(* CODESYS project Example8_PLC.project

Project tree, tasks and I/O mapping:
  Device : CODESYS Control Win V3, 3S - Smart Software Solutions GmbH, order no. 305021, version 3.5.7.0
    application Application
      libraries: Standard, * (System)
      task MainTask (cyclic, interval t#20ms, priority 1) calls PLC_PRG
      program PLC_PRG [ST]
      global variables GVL
      function block FB_G4LTL [ST]
    Ethernet : Ethernet, 3S - Smart Software Solutions GmbH, version 3.5.7.0
      Modbus_TCP_Master : Modbus TCP Master, 3S - Smart Software Solutions GmbH, version 3.5.6.0
          settings: AutoReconnect = TRUE
        Modbus_TCP_Slave : Modbus TCP Slave, 3S - Smart Software Solutions GmbH, version 3.5.7.0
            settings: Unit-ID = 1; IPAddress = [127, 0, 0, 1]; Channel 0.Function Code = 4; Channel 0.Read Offset = 16#0000; Channel 0.Read Length = 1; Channel 0.Write Offset = 0; Channel 0.Write Length = 0; Channel 0.Cycle Time = 100; Channel 1.Function Code = 4; Channel 1.Read Offset = 16#0001; Channel 1.Read Length = 1; Channel 1.Write Offset = 0; Channel 1.Write Length = 0; Channel 1.Cycle Time = 100; Channel 2.Function Code = 4; Channel 2.Read Offset = 16#0002; Channel 2.Read Length = 1; Channel 2.Write Offset = 0; Channel 2.Write Length = 0; Channel 2.Cycle Time = 100; Channel 3.Function Code = 4; Channel 3.Read Offset = 16#0003; Channel 3.Read Length = 1; Channel 3.Write Offset = 0; Channel 3.Write Length = 0; Channel 3.Cycle Time = 100; Channel 4.Function Code = 4; Channel 4.Read Offset = 16#0004; Channel 4.Read Length = 1; Channel 4.Write Offset = 0; Channel 4.Write Length = 0; Channel 4.Cycle Time = 100; Channel 5.Function Code = 6; Channel 5.Read Offset = 0; Channel 5.Read Length = 0; Channel 5.Write Offset = 16#0000; Channel 5.Write Length = 1; Channel 5.Cycle Time = 100; Channel 6.Function Code = 6; Channel 6.Read Offset = 0;
              Channel 6.Read Length = 0; Channel 6.Write Offset = 16#0002; Channel 6.Write Length = 1; Channel 6.Cycle Time = 100; Channel 7.Function Code = 6; Channel 7.Read Offset = 0; Channel 7.Read Length = 0; Channel 7.Write Offset = 16#0003; Channel 7.Write Length = 1; Channel 7.Cycle Time = 100; Channel 8.Function Code = 6; Channel 8.Read Offset = 0; Channel 8.Read Length = 0; Channel 8.Write Offset = 16#0004; Channel 8.Write Length = 1; Channel 8.Cycle Time = 100; Channel 9.Function Code = 6; Channel 9.Read Offset = 0; Channel 9.Read Length = 0; Channel 9.Write Offset = 16#0001; Channel 9.Write Length = 1; Channel 9.Cycle Time = 100
            input  Application.dIn0 : BOOL  // Channel 0.Channel 0.Bit0
            input  Application.dIn1 : BOOL  // Channel 1.Channel 1.Bit0
            input  Application.dIn2 : BOOL  // Channel 2.Channel 2.Bit0
            input  Application.dIn3 : BOOL  // Channel 3.Channel 3.Bit0
            input  Application.dIn4 : BOOL  // Channel 4.Channel 4.Bit0
            output Application.dOut0 : BOOL  // Channel 5.Channel 5.Bit0
            output Application.dOut2 : BOOL  // Channel 6.Channel 6.Bit0
            output Application.dOut3 : BOOL  // Channel 7.Channel 7.Bit0
            output Application.dOut4 : BOOL  // Channel 8.Channel 8.Bit0
            output Application.dOut1 : BOOL  // Channel 9.Channel 9.Bit0
            unmapped channels: Channel 0, Channel 1, Channel 2, Channel 3, Channel 4, Channel 5, Channel 6, Channel 7, Channel 8, Channel 9
*)

// Device/Application/GVL
VAR_GLOBAL
	
dIn0 : BOOL;
dIn1 : BOOL;
dIn2 : BOOL;
dIn3 : BOOL;
dIn4 : BOOL;

dOut0 : BOOL;
dOut1 : BOOL; 
dOut2 : BOOL; 
dOut3 : BOOL; 
dOut4 : BOOL; 
END_VAR

// Device/Application/PLC_PRG
PROGRAM PLC_PRG

VAR 
	fb: FB_G4LTL;
END_VAR


// Direct looping
// Assign pins (from global variable to function block) 
fb.x1 := dIn0;

// Assign pins (from function block to global variable)
dOut0 := fb.y1;

// Run the function block
fb();

END_PROGRAM

// Device/Application/FB_G4LTL
FUNCTION_BLOCK FB_G4LTL
 
   (* Variable definition *)
   VAR_INPUT
      x1	: BOOL;
   END_VAR
   VAR_OUTPUT
      y1	: BOOL;
   END_VAR
   VAR
   (* The total number of states equals to 7 *)
      cstate86	: LINT := 0;
      t0	: TON;
      t0_reset	: BOOL := FALSE;
      t0_up	: BOOL := FALSE;
      t0_start	: BOOL := FALSE;
	  
      t1	: TON;
      t1_reset	: BOOL := FALSE;
      t1_up	: BOOL := FALSE;
      t1_start	: BOOL := FALSE;
	  
	  T0_VALUE	: TIME := TIME#5S;
      T1_VALUE	: TIME := TIME#3s;
	  
   END_VAR

   (* Constant definition (depending on compiler, one might need to move to normal variables) *)

   (* Control logic *)
CASE cstate86 OF
424082:
    IF ((x1 = FALSE) AND  ( TRUE ) AND  (t1.Q = FALSE)) THEN 
        cstate86 := 924337; y1 := TRUE; t0_start := FALSE;t1_start := TRUE; t1_up := FALSE; 
    ELSIF ((x1 = FALSE) AND  ( TRUE ) AND  (t1.Q = TRUE)) THEN 
        cstate86 := 924341; y1 := TRUE; t0_start := FALSE;t1_start := TRUE; t1_up := FALSE; 
    ELSIF ((x1 = TRUE) AND  (t0.Q = FALSE) AND  ( TRUE )) THEN 
        cstate86 := 403602; y1 := FALSE; t0_start := FALSE;t1_start := FALSE; 
    ELSIF ((x1 = TRUE) AND  (t0.Q = TRUE) AND  ( TRUE )) THEN 
        cstate86 := 424082; y1 := TRUE; t0_start := FALSE;t1_start := FALSE; 
    END_IF;
270866:
    IF ((x1 = FALSE) AND  ( TRUE ) AND  (t1.Q = FALSE)) THEN 
        cstate86 := 993810; y1 := FALSE; t0_start := FALSE;t1_start := FALSE; 
    ELSIF ((x1 = FALSE) AND  ( TRUE ) AND  (t1.Q = TRUE)) THEN 
        cstate86 := 993048; y1 := FALSE; t0_start := FALSE;t1_start := FALSE; 
    ELSIF ((x1 = TRUE) AND  (t0.Q = FALSE) AND  ( TRUE )) THEN 
        cstate86 := 543012; y1 := FALSE; t0_start := TRUE; t0_up := FALSE;t1_start := FALSE; 
    ELSIF ((x1 = TRUE) AND  (t0.Q = TRUE) AND  ( TRUE )) THEN 
        cstate86 := 551204; y1 := FALSE; t0_start := TRUE; t0_up := FALSE;t1_start := FALSE; 
    END_IF;
403602:
    IF ((x1 = FALSE) AND  ( TRUE ) AND  (t1.Q = FALSE)) THEN 
        cstate86 := 924337; y1 := TRUE; t0_start := FALSE;t1_start := TRUE; t1_up := FALSE; 
    ELSIF ((x1 = FALSE) AND  ( TRUE ) AND  (t1.Q = TRUE)) THEN 
        cstate86 := 924341; y1 := TRUE; t0_start := FALSE;t1_start := TRUE; t1_up := FALSE; 
    ELSIF ((x1 = TRUE) AND  (t0.Q = FALSE) AND  ( TRUE )) THEN 
        cstate86 := 403602; y1 := FALSE; t0_start := FALSE;t1_start := FALSE; 
    ELSIF ((x1 = TRUE) AND  (t0.Q = TRUE) AND  ( TRUE )) THEN 
        cstate86 := 424082; y1 := FALSE; t0_start := FALSE;t1_start := FALSE; 
    END_IF;
270872:
    IF ((x1 = FALSE) AND  ( TRUE ) AND  (t1.Q = FALSE)) THEN 
        cstate86 := 993810; y1 := FALSE; t0_start := FALSE;t1_start := FALSE; 
    ELSIF ((x1 = FALSE) AND  ( TRUE ) AND  (t1.Q = TRUE)) THEN 
        cstate86 := 993048; y1 := FALSE; t0_start := FALSE;t1_start := FALSE; 
    ELSIF ((x1 = TRUE) AND  (t0.Q = FALSE) AND  ( TRUE )) THEN 
        cstate86 := 543012; y1 := FALSE; t0_start := TRUE; t0_up := FALSE;t1_start := FALSE; 
    ELSIF ((x1 = TRUE) AND  (t0.Q = TRUE) AND  ( TRUE )) THEN 
        cstate86 := 551204; y1 := FALSE; t0_start := TRUE; t0_up := FALSE;t1_start := FALSE; 
    END_IF;
993048:
    IF ((x1 = FALSE) AND  ( TRUE ) AND  (t1.Q = FALSE)) THEN 
        cstate86 := 993810; y1 := FALSE; t0_start := FALSE;t1_start := FALSE; 
    ELSIF ((x1 = FALSE) AND  ( TRUE ) AND  (t1.Q = TRUE)) THEN 
        cstate86 := 993048; y1 := FALSE; t0_start := FALSE;t1_start := FALSE; 
    ELSIF ((x1 = TRUE) AND  (t0.Q = FALSE) AND  ( TRUE )) THEN 
        cstate86 := 543012; y1 := FALSE; t0_start := TRUE; t0_up := FALSE;t1_start := FALSE; 
    ELSIF ((x1 = TRUE) AND  (t0.Q = TRUE) AND  ( TRUE )) THEN 
        cstate86 := 551204; y1 := FALSE; t0_start := TRUE; t0_up := FALSE;t1_start := FALSE; 
    END_IF;
551204:
    IF ((x1 = FALSE) AND  (t0.Q = FALSE) AND  ( TRUE )) THEN 
        cstate86 := 697833; y1 := FALSE; t0_start := FALSE;t1_start := FALSE; 
    ELSIF ((x1 = FALSE) AND  (t0.Q = TRUE) AND  (t1.Q = FALSE)) THEN 
        cstate86 := 924337; y1 := TRUE; t0_start := FALSE;t1_start := TRUE; t1_up := FALSE; 
    ELSIF ((x1 = FALSE) AND  (t0.Q = TRUE) AND  (t1.Q = TRUE)) THEN 
        cstate86 := 924341; y1 := TRUE; t0_start := FALSE;t1_start := TRUE; t1_up := FALSE; 
    ELSIF ((x1 = TRUE) AND  (t0.Q = FALSE) AND  ( TRUE )) THEN 
        cstate86 := 870436; y1 := FALSE; t0_start := FALSE;t1_start := FALSE; 
    ELSIF ((x1 = TRUE) AND  (t0.Q = TRUE) AND  ( TRUE )) THEN 
        cstate86 := 423570; y1 := TRUE; t0_start := FALSE;t1_start := FALSE; 
    END_IF;
422674:
    IF ((x1 = FALSE) AND  ( TRUE ) AND  (t1.Q = FALSE)) THEN 
        cstate86 := 924337; y1 := TRUE; t0_start := FALSE;t1_start := TRUE; t1_up := FALSE; 
    ELSIF ((x1 = FALSE) AND  ( TRUE ) AND  (t1.Q = TRUE)) THEN 
        cstate86 := 924341; y1 := TRUE; t0_start := FALSE;t1_start := TRUE; t1_up := FALSE; 
    ELSIF ((x1 = TRUE) AND  (t0.Q = FALSE) AND  ( TRUE )) THEN 
        cstate86 := 403602; y1 := FALSE; t0_start := FALSE;t1_start := FALSE; 
    ELSIF ((x1 = TRUE) AND  (t0.Q = TRUE) AND  ( TRUE )) THEN 
        cstate86 := 424082; y1 := TRUE; t0_start := FALSE;t1_start := FALSE; 
    END_IF;
697833:
    IF (( true )) THEN 
        cstate86 := 697833; y1 := FALSE; t0_start := FALSE;t1_start := FALSE; 
    END_IF;
870436:
    IF ((x1 = FALSE) AND  (t0.Q = FALSE) AND  ( TRUE )) THEN 
        cstate86 := 697833; y1 := FALSE; t0_start := FALSE;t1_start := FALSE; 
    ELSIF ((x1 = FALSE) AND  (t0.Q = TRUE) AND  (t1.Q = FALSE)) THEN 
        cstate86 := 924337; y1 := TRUE; t0_start := FALSE;t1_start := TRUE; t1_up := FALSE; 
    ELSIF ((x1 = FALSE) AND  (t0.Q = TRUE) AND  (t1.Q = TRUE)) THEN 
        cstate86 := 924341; y1 := TRUE; t0_start := FALSE;t1_start := TRUE; t1_up := FALSE; 
    ELSIF ((x1 = TRUE) AND  (t0.Q = FALSE) AND  ( TRUE )) THEN 
        cstate86 := 870436; y1 := FALSE; t0_start := FALSE;t1_start := FALSE; 
    ELSIF ((x1 = TRUE) AND  (t0.Q = TRUE) AND  ( TRUE )) THEN 
        cstate86 := 423570; y1 := FALSE; t0_start := FALSE;t1_start := FALSE; 
    END_IF;
402194:
    IF ((x1 = FALSE) AND  ( TRUE ) AND  (t1.Q = FALSE)) THEN 
        cstate86 := 924337; y1 := TRUE; t0_start := FALSE;t1_start := TRUE; t1_up := FALSE; 
    ELSIF ((x1 = FALSE) AND  ( TRUE ) AND  (t1.Q = TRUE)) THEN 
        cstate86 := 924341; y1 := TRUE; t0_start := FALSE;t1_start := TRUE; t1_up := FALSE; 
    ELSIF ((x1 = TRUE) AND  (t0.Q = FALSE) AND  ( TRUE )) THEN 
        cstate86 := 403602; y1 := FALSE; t0_start := FALSE;t1_start := FALSE; 
    ELSIF ((x1 = TRUE) AND  (t0.Q = TRUE) AND  ( TRUE )) THEN 
        cstate86 := 424082; y1 := FALSE; t0_start := FALSE;t1_start := FALSE; 
    END_IF;
0:
    IF ((x1 = FALSE) AND  ( TRUE ) AND  (t1.Q = FALSE)) THEN 
        cstate86 := 270866; y1 := FALSE; t0_start := FALSE;t1_start := FALSE; 
    ELSIF ((x1 = FALSE) AND  ( TRUE ) AND  (t1.Q = TRUE)) THEN 
        cstate86 := 270872; y1 := FALSE; t0_start := FALSE;t1_start := FALSE; 
    ELSIF ((x1 = TRUE) AND  (t0.Q = FALSE) AND  ( TRUE )) THEN 
        cstate86 := 402194; y1 := FALSE; t0_start := FALSE;t1_start := FALSE; 
    ELSIF ((x1 = TRUE) AND  (t0.Q = TRUE) AND  ( TRUE )) THEN 
        cstate86 := 422674; y1 := FALSE; t0_start := FALSE;t1_start := FALSE; 
    END_IF;
423570:
    IF ((x1 = FALSE) AND  ( TRUE ) AND  (t1.Q = FALSE)) THEN 
        cstate86 := 924337; y1 := TRUE; t0_start := FALSE;t1_start := TRUE; t1_up := FALSE; 
    ELSIF ((x1 = FALSE) AND  ( TRUE ) AND  (t1.Q = TRUE)) THEN 
        cstate86 := 924341; y1 := TRUE; t0_start := FALSE;t1_start := TRUE; t1_up := FALSE; 
    ELSIF ((x1 = TRUE) AND  (t0.Q = FALSE) AND  ( TRUE )) THEN 
        cstate86 := 403602; y1 := FALSE; t0_start := FALSE;t1_start := FALSE; 
    ELSIF ((x1 = TRUE) AND  (t0.Q = TRUE) AND  ( TRUE )) THEN 
        cstate86 := 424082; y1 := TRUE; t0_start := FALSE;t1_start := FALSE; 
    END_IF;
924337:
    IF ((x1 = FALSE) AND  ( TRUE ) AND  (t1.Q = FALSE)) THEN 
        cstate86 := 595121; y1 := TRUE; t0_start := FALSE;t1_start := FALSE; 
    ELSIF ((x1 = FALSE) AND  ( TRUE ) AND  (t1.Q = TRUE)) THEN 
        cstate86 := 730904; y1 := FALSE; t0_start := FALSE;t1_start := FALSE; 
    ELSIF ((x1 = TRUE) AND  ( TRUE ) AND  (t1.Q = FALSE)) THEN 
        cstate86 := 697833; y1 := FALSE; t0_start := FALSE;t1_start := FALSE; 
    ELSIF ((x1 = TRUE) AND  (t0.Q = FALSE) AND  (t1.Q = TRUE)) THEN 
        cstate86 := 543012; y1 := FALSE; t0_start := TRUE; t0_up := FALSE;t1_start := FALSE; 
    ELSIF ((x1 = TRUE) AND  (t0.Q = TRUE) AND  (t1.Q = TRUE)) THEN 
        cstate86 := 551204; y1 := FALSE; t0_start := TRUE; t0_up := FALSE;t1_start := FALSE; 
    END_IF;
993810:
    IF ((x1 = FALSE) AND  ( TRUE ) AND  (t1.Q = FALSE)) THEN 
        cstate86 := 993810; y1 := FALSE; t0_start := FALSE;t1_start := FALSE; 
    ELSIF ((x1 = FALSE) AND  ( TRUE ) AND  (t1.Q = TRUE)) THEN 
        cstate86 := 993048; y1 := FALSE; t0_start := FALSE;t1_start := FALSE; 
    ELSIF ((x1 = TRUE) AND  (t0.Q = FALSE) AND  ( TRUE )) THEN 
        cstate86 := 543012; y1 := FALSE; t0_start := TRUE; t0_up := FALSE;t1_start := FALSE; 
    ELSIF ((x1 = TRUE) AND  (t0.Q = TRUE) AND  ( TRUE )) THEN 
        cstate86 := 551204; y1 := FALSE; t0_start := TRUE; t0_up := FALSE;t1_start := FALSE; 
    END_IF;
595121:
    IF ((x1 = FALSE) AND  ( TRUE ) AND  (t1.Q = FALSE)) THEN 
        cstate86 := 595121; y1 := TRUE; t0_start := FALSE;t1_start := FALSE; 
    ELSIF ((x1 = FALSE) AND  ( TRUE ) AND  (t1.Q = TRUE)) THEN 
        cstate86 := 730904; y1 := FALSE; t0_start := FALSE;t1_start := FALSE; 
    ELSIF ((x1 = TRUE) AND  ( TRUE ) AND  (t1.Q = FALSE)) THEN 
        cstate86 := 697833; y1 := FALSE; t0_start := FALSE;t1_start := FALSE; 
    ELSIF ((x1 = TRUE) AND  (t0.Q = FALSE) AND  (t1.Q = TRUE)) THEN 
        cstate86 := 543012; y1 := FALSE; t0_start := TRUE; t0_up := FALSE;t1_start := FALSE; 
    ELSIF ((x1 = TRUE) AND  (t0.Q = TRUE) AND  (t1.Q = TRUE)) THEN 
        cstate86 := 551204; y1 := FALSE; t0_start := TRUE; t0_up := FALSE;t1_start := FALSE; 
    END_IF;
543012:
    IF ((x1 = FALSE) AND  (t0.Q = FALSE) AND  ( TRUE )) THEN 
        cstate86 := 697833; y1 := FALSE; t0_start := FALSE;t1_start := FALSE; 
    ELSIF ((x1 = FALSE) AND  (t0.Q = TRUE) AND  (t1.Q = FALSE)) THEN 
        cstate86 := 924337; y1 := TRUE; t0_start := FALSE;t1_start := TRUE; t1_up := FALSE; 
    ELSIF ((x1 = FALSE) AND  (t0.Q = TRUE) AND  (t1.Q = TRUE)) THEN 
        cstate86 := 924341; y1 := TRUE; t0_start := FALSE;t1_start := TRUE; t1_up := FALSE; 
    ELSIF ((x1 = TRUE) AND  (t0.Q = FALSE) AND  ( TRUE )) THEN 
        cstate86 := 870436; y1 := FALSE; t0_start := FALSE;t1_start := FALSE; 
    ELSIF ((x1 = TRUE) AND  (t0.Q = TRUE) AND  ( TRUE )) THEN 
        cstate86 := 423570; y1 := FALSE; t0_start := FALSE;t1_start := FALSE; 
    END_IF;
924341:
    IF ((x1 = FALSE) AND  ( TRUE ) AND  (t1.Q = FALSE)) THEN 
        cstate86 := 595121; y1 := TRUE; t0_start := FALSE;t1_start := FALSE; 
    ELSIF ((x1 = FALSE) AND  ( TRUE ) AND  (t1.Q = TRUE)) THEN 
        cstate86 := 730904; y1 := FALSE; t0_start := FALSE;t1_start := FALSE; 
    ELSIF ((x1 = TRUE) AND  ( TRUE ) AND  (t1.Q = FALSE)) THEN 
        cstate86 := 697833; y1 := FALSE; t0_start := FALSE;t1_start := FALSE; 
    ELSIF ((x1 = TRUE) AND  (t0.Q = FALSE) AND  (t1.Q = TRUE)) THEN 
        cstate86 := 543012; y1 := FALSE; t0_start := TRUE; t0_up := FALSE;t1_start := FALSE; 
    ELSIF ((x1 = TRUE) AND  (t0.Q = TRUE) AND  (t1.Q = TRUE)) THEN 
        cstate86 := 551204; y1 := FALSE; t0_start := TRUE; t0_up := FALSE;t1_start := FALSE; 
    END_IF;
730904:
    IF ((x1 = FALSE) AND  ( TRUE ) AND  (t1.Q = FALSE)) THEN 
        cstate86 := 993810; y1 := FALSE; t0_start := FALSE;t1_start := FALSE; 
    ELSIF ((x1 = FALSE) AND  ( TRUE ) AND  (t1.Q = TRUE)) THEN 
        cstate86 := 993048; y1 := FALSE; t0_start := FALSE;t1_start := FALSE; 
    ELSIF ((x1 = TRUE) AND  (t0.Q = FALSE) AND  ( TRUE )) THEN 
        cstate86 := 543012; y1 := FALSE; t0_start := TRUE; t0_up := FALSE;t1_start := FALSE; 
    ELSIF ((x1 = TRUE) AND  (t0.Q = TRUE) AND  ( TRUE )) THEN 
        cstate86 := 551204; y1 := FALSE; t0_start := TRUE; t0_up := FALSE;t1_start := FALSE; 
    END_IF;
END_CASE;

(* Additional processing to handle clocks - in CODESYS, it only starts
    with rising edge and can not be placed inside IF statement *) 
IF(t0_up = TRUE) THEN
    t0_reset := TRUE;
ELSIF(t0_start = TRUE AND t0_up = FALSE) THEN
    t0_up := TRUE;  t0_reset := FALSE;
END_IF
t0(IN:=t0_reset, PT:=T0_VALUE); 
IF(t1_up = TRUE) THEN
    t1_reset := TRUE;
ELSIF(t1_start = TRUE AND t1_up = FALSE) THEN
    t1_up := TRUE;  t1_reset := FALSE;
END_IF
t1(IN:=t1_reset, PT:=T1_VALUE);

END_FUNCTION_BLOCK
